// TwinCAT 3 PLC project IO_ReadWrite
// Title: IO_ReadWrite
// Company: BACA_Apps
// ProjectVersion: 0.0.0.1
// ProgramVersion: 3.1.4026.27
// libraries:
//   Tc2_Standard, * (Beckhoff Automation GmbH)
//   Tc2_System, * (Beckhoff Automation GmbH)
// project tree:
//   POUs/ FB_IO_ReadWrite.TcPOU
// real-time tasks:
//   TASK PlcTask1: cycle T#1ms, priority 21, ADS port 351
// I/O:
//   DEVICE Device 1 (EtherCAT), AmsNetId 5.143.132.242.2.1
//     Term 1 (EK1200) [EK1200-5000 EtherCAT Power supply (2A E-Bus)]
//       Term 2 (EL1002) [EL1002 2Ch. Dig. Input 24V, 3ms]
//       Term 3 (EL2002) [EL2002 2Ch. Dig. Output 24V, 0.5A]
//       Term 4 (EL9011) [EL9011 End Terminal]
// variable links:
//   TestFrameworkPLC/TestFrameworkPLC Instance <-> Device 1 (EtherCAT)/Term 1 (EK1200)/Term 2 (EL1002)
//     PlcTask Inputs/MAIN.fbT1.fbIOtester.bIn <-> Channel 1/Input
//   TestFrameworkPLC/TestFrameworkPLC Instance <-> Device 1 (EtherCAT)/Term 1 (EK1200)/Term 3 (EL2002)
//     PlcTask Outputs/MAIN.fbT1.fbIOtester.bOut <-> Channel 1/Output

// ---- POUs/FB_IO_ReadWrite.TcPOU
{ attribute 'Name' := 'TC_DI-DO-Test' }
{ attribute 'Timeout' := 't#5s' }
{ attribute 'Owner' := 'BACA_Controls' }
{ attribute 'Category' := 'IO/Digital' }
FUNCTION_BLOCK FB_IO_ReadWrite
VAR_INPUT
	bExecute     : BOOL;           
	timerDelay   : TIME; 
END_VAR
VAR_OUTPUT
	bHighMatch   : BOOL;           
	bLowMatch    : BOOL;   
	bDone 		 : BOOL;        
END_VAR
VAR
	rTrigExecute : R_TRIG;
	bOut AT %Q*	 : BOOL;
	bIn  AT %I*  : BOOL;
	timer        : TON;
	eState       : (INIT, SET_TRUE, READ_TRUE, SET_FALSE, READ_FALSE);
END_VAR

rTrigExecute(CLK := bExecute);

CASE eState OF
	INIT:
		bOut := FALSE;
		bHighMatch := FALSE;
		bLowMatch := FALSE;
		bDone := FALSE;
		timer.PT := timerDelay;
		IF rTrigExecute.Q THEN
			eState := SET_TRUE;
		END_IF

	SET_TRUE:
		bOut := TRUE;
		timer.IN := TRUE;
		IF timer.Q THEN
			timer.IN := FALSE;
			eState := READ_TRUE;
		END_IF;

	READ_TRUE:
		bHighMatch := (bIn = TRUE);		
		eState := SET_FALSE;

	SET_FALSE:
		bOut := FALSE;
		timer.IN := TRUE;
		IF timer.Q THEN
			timer.IN := FALSE;
			eState := READ_FALSE;
		END_IF;

	READ_FALSE:
		bLowMatch := (bIn = FALSE);
		bDone := TRUE;
		eState := INIT;
END_CASE

timer();

END_FUNCTION_BLOCK
